// TIA Portal V20 export
VAR_GLOBAL   // PLC tag table "Safety"
   "IS_NOT-HALT_Taster_1_Kanal_A" AT %I100.0 : Bool;   // IS +Feld=EAS-131S1 NOT-HALT Taster 1, Kanal A
   "IS_NOT-HALT_Extern_2_Kanal_A" AT %I100.2 : Bool;   // IS + __________ NOT-HALT Extern 2, Kanal A
   IS_Tuer_1_Kanal_A AT %I100.4 : Bool;   // IS +Feld=STÜR-921S1/S2 Tür 1, Kanal A
   IS_Tuer_2_Kanal_A AT %I100.5 : Bool;   // IS +___________ Tür 2 oder Lichtvorhang, Kanal A
   "IS_NOT-HALT_Taster_1_Kanal_B" AT %I101.0 : Bool;   // IS +Feld=EAS-131S1 NOT-HALT Taster 1, Kanal B
   "IS_NOT-HALT_Extern_1_Kanal_B" AT %I101.1 : Bool;   // IS +HS1=ÜSPS-125K1/K2 NOT-HALT Extern 1, Kanal B
   "IS_NOT-HALT_Extern_2_Kanal_B" AT %I101.2 : Bool;   // IS +___________ NOT-HALT Extern 2, Kanal B
   "IS_NOT-HALT_Extern_1_Kanal_A" AT %I100.1 : Bool;   // IS +HS1=ÜSPS-125K1/K2 NOT-HALT Extern 1, Kanal A
   "QS_NOT-HALT_Schuetz" AT %Q110.0 : Bool;   // QS +HS1=AAS-146K1 NOT-HALT Schütz
   "QS_NOT-HALT_Tuere_1_RST" AT %Q110.1 : Bool;   // QS +_______ NOT-HALT Türe 1 RST
   "QS_NOT-HALT_Tuere_2_RST" AT %Q110.3 : Bool;   // QS +_______ NOT-HALT Türe 2 RST
   "QS_NOT-HALT_Tuere_2" AT %Q110.4 : Bool;   // QS +_______ NOT-HALT Türe 2
   "QS_NOT-HALT_Roboter" AT %Q110.5 : Bool;   // QS +_______ NOT-HALT Roboter
   QS_Sichere_Bewegung AT %Q110.6 : Bool;   // QS +_______ Sichere Bewegung
   "QS_NOT-HALT_Tuere_1" AT %Q110.2 : Bool;   // QS +HS1=AAS-148K1 NOT-HALT Türe 1
   IS_Tuer_1_Kanal_B AT %I101.4 : Bool;   // IS +Feld=STÜR-921S1/S2 Tür 1, Kanal B
   IS_Tuer_2_Kanal_B AT %I101.5 : Bool;   // IS +___________ Tür 2 oder Lichtvorhang, Kanal B
   IS_Zustimmtaster_Kanal_A AT %I100.3 : Bool;   // IS +HS1=ÜSPS-125K1/K2 Zustimmtaster, Kanal A
   IS_Rueck_Entlueftung AT %I100.6 : Bool;   // IS +___________ Rück Entlüftet
   IS_Druckbereich_entlueftet AT %I100.7 : Bool;   // IS +Feld=PV-938S2 Druckbereich entlüftet
   IS_Zustimmtaster_Kanal_B AT %I101.3 : Bool;   // IS +HS1=ÜSPS-125K1/K2 Zustimmtaster, Kanal B
   IS_Systemdruck_OK AT %I101.6 : Bool;   // IS +Feld=PV-938S1 Systemdruck OK
   IS101_7 AT %I101.7 : Bool;
   QS_Zuhaltung_Freigeben AT %Q110.7 : Bool;   // QS +HS1=AAS-151K1 Zuhaltung Freigeben
END_VAR
